// Mitsubishi GX Works2 project: AGV_IOCHECK   PLC: Q03UD

PROGRAM IOCHECK
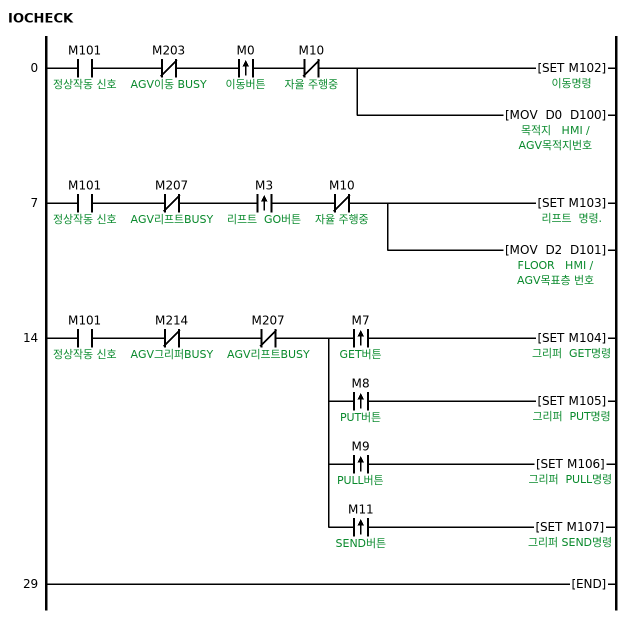
0     LD      M101  ; 정상작동 신호
      ANI     M203  ; AGV이동 BUSY
      ANDP    M0  ; 이동버튼
      ANI     M10  ; 자율 주행중
      SET     M102  ; 이동명령
      MOV     D0 D100  ; 목적지   HMI / AGV목적지번호
7     LD      M101  ; 정상작동 신호
      ANI     M207  ; AGV리프트BUSY
      ANDP    M3  ; 리프트  GO버튼
      ANI     M10  ; 자율 주행중
      SET     M103  ; 리프트  명령.
      MOV     D2 D101  ; FLOOR   HMI / AGV목표층 번호
14    LD      M101  ; 정상작동 신호
      ANI     M214  ; AGV그리퍼BUSY
      ANI     M207  ; AGV리프트BUSY
      MPS
      ANDP    M7  ; GET버튼
      SET     M104  ; 그리퍼  GET명령
      MRD
      ANDP    M8  ; PUT버튼
      SET     M105  ; 그리퍼  PUT명령
      MRD
      ANDP    M9  ; PULL버튼
      SET     M106  ; 그리퍼  PULL명령
      MPP
      ANDP    M11  ; SEND버튼
      SET     M107  ; 그리퍼 SEND명령
29    END
END_PROGRAM

PROGRAM MAIN
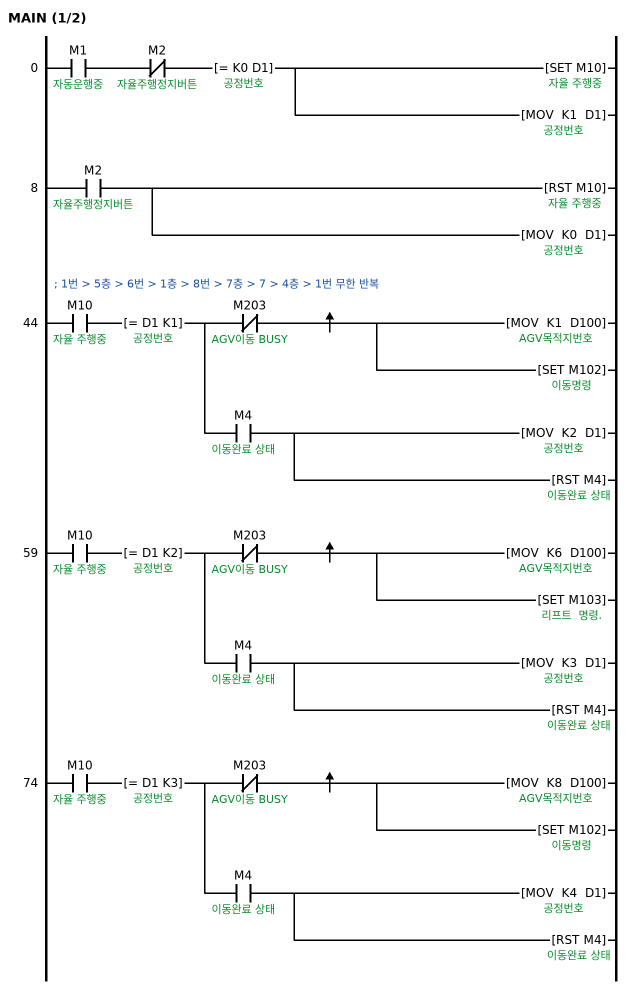
0     LD      M1  ; 자동운행중
      ANI     M2  ; 자율주행정지버튼
      AND=    K0 D1  ; 공정번호
      SET     M10  ; 자율 주행중
      MOV     K1 D1
8     LD      M2  ; 자율주행정지버튼
      RST     M10  ; 자율 주행중
      MOV     K0 D1
; 1번 > 5층 > 6번 > 1층 > 8번 > 7층 > 7 > 4층 > 1번 무한 반복
44    LD      M10  ; 자율 주행중
      AND=    D1 K1  ; 공정번호
      MPS
      ANI     M203  ; AGV이동 BUSY
      MEP
      MOV     K1 D100  ; AGV목적지번호
      SET     M102  ; 이동명령
      MPP
      AND     M4  ; 이동완료 상태
      MOV     K2 D1
      RST     M4  ; 이동완료 상태
59    LD      M10  ; 자율 주행중
      AND=    D1 K2  ; 공정번호
      MPS
      ANI     M203  ; AGV이동 BUSY
      MEP
      MOV     K6 D100
      SET     M103  ; 리프트  명령.
      MPP
      AND     M4  ; 이동완료 상태
      MOV     K3 D1
      RST     M4  ; 이동완료 상태
74    LD      M10  ; 자율 주행중
      AND=    D1 K3  ; 공정번호
      MPS
      ANI     M203  ; AGV이동 BUSY
      MEP
      MOV     K8 D100
      SET     M102  ; 이동명령
      MPP
      AND     M4  ; 이동완료 상태
      MOV     K4 D1
      RST     M4  ; 이동완료 상태
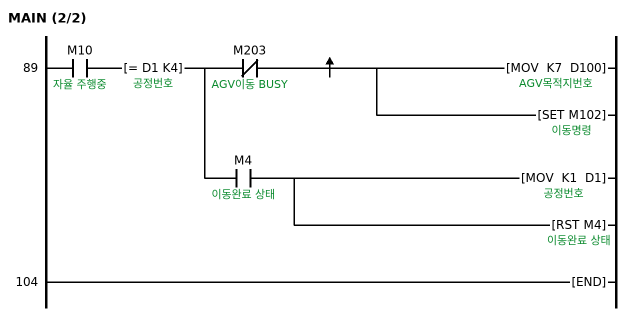
89    LD      M10  ; 자율 주행중
      AND=    D1 K4  ; 공정번호
      MPS
      ANI     M203  ; AGV이동 BUSY
      MEP
      MOV     K7 D100
      SET     M102  ; 이동명령
      MPP
      AND     M4  ; 이동완료 상태
      MOV     K1 D1
      RST     M4  ; 이동완료 상태
104   END
END_PROGRAM

PROGRAM MAIN2
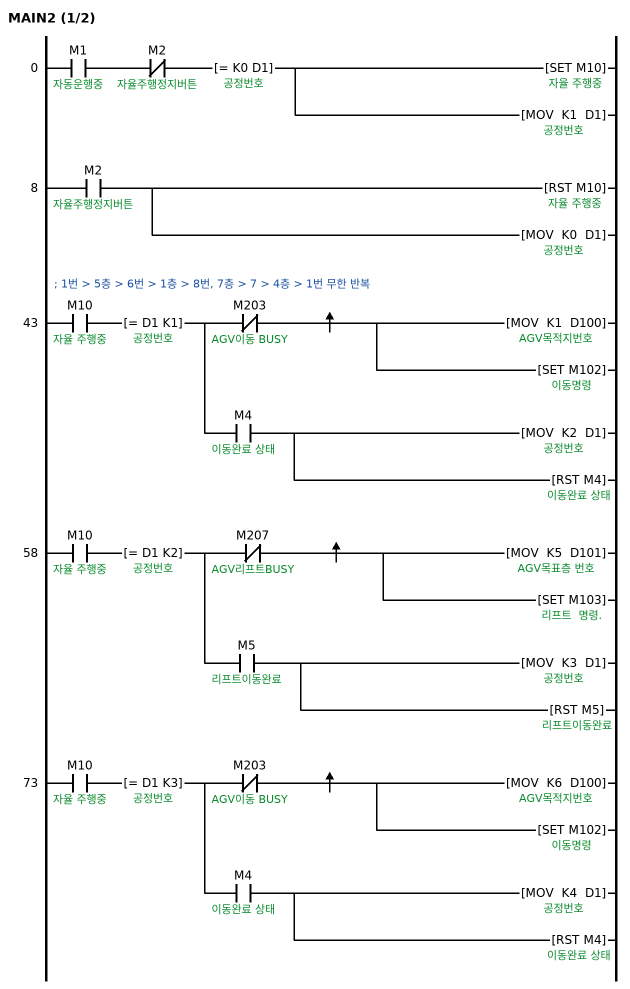
0     LD      M1  ; 자동운행중
      ANI     M2  ; 자율주행정지버튼
      AND=    K0 D1  ; 공정번호
      SET     M10  ; 자율 주행중
      MOV     K1 D1
8     LD      M2  ; 자율주행정지버튼
      RST     M10  ; 자율 주행중
      MOV     K0 D1
; 1번 > 5층 > 6번 > 1층 > 8번, 7층 > 7 > 4층 > 1번 무한 반복
43    LD      M10  ; 자율 주행중
      AND=    D1 K1  ; 공정번호
      MPS
      ANI     M203  ; AGV이동 BUSY
      MEP
      MOV     K1 D100  ; AGV목적지번호
      SET     M102  ; 이동명령
      MPP
      AND     M4  ; 이동완료 상태
      MOV     K2 D1
      RST     M4  ; 이동완료 상태
58    LD      M10  ; 자율 주행중
      AND=    D1 K2  ; 공정번호
      MPS
      ANI     M207  ; AGV리프트BUSY
      MEP
      MOV     K5 D101  ; AGV목표층 번호
      SET     M103  ; 리프트  명령.
      MPP
      AND     M5  ; 리프트이동완료
      MOV     K3 D1
      RST     M5  ; 리프트이동완료
73    LD      M10  ; 자율 주행중
      AND=    D1 K3  ; 공정번호
      MPS
      ANI     M203  ; AGV이동 BUSY
      MEP
      MOV     K6 D100
      SET     M102  ; 이동명령
      MPP
      AND     M4  ; 이동완료 상태
      MOV     K4 D1
      RST     M4  ; 이동완료 상태
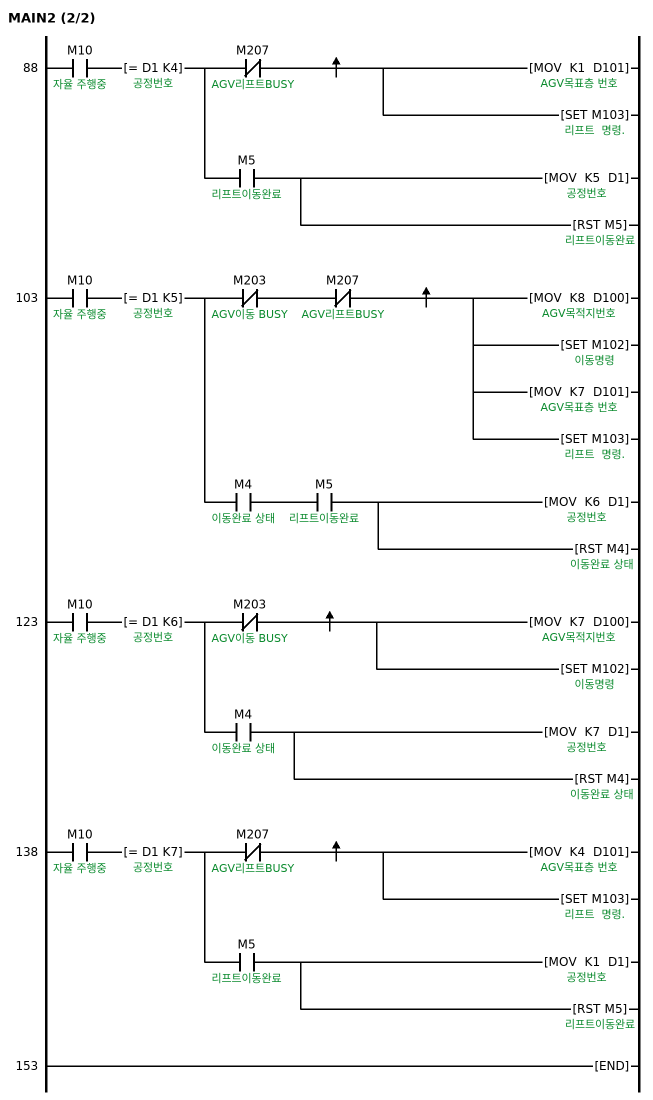
88    LD      M10  ; 자율 주행중
      AND=    D1 K4  ; 공정번호
      MPS
      ANI     M207  ; AGV리프트BUSY
      MEP
      MOV     K1 D101
      SET     M103  ; 리프트  명령.
      MPP
      AND     M5  ; 리프트이동완료
      MOV     K5 D1
      RST     M5  ; 리프트이동완료
103   LD      M10  ; 자율 주행중
      AND=    D1 K5  ; 공정번호
      MPS
      ANI     M203  ; AGV이동 BUSY
      ANI     M207  ; AGV리프트BUSY
      MEP
      MOV     K8 D100
      SET     M102  ; 이동명령
      MOV     K7 D101
      SET     M103  ; 리프트  명령.
      MPP
      AND     M4  ; 이동완료 상태
      AND     M5  ; 리프트이동완료
      MOV     K6 D1
      RST     M4  ; 이동완료 상태
123   LD      M10  ; 자율 주행중
      AND=    D1 K6  ; 공정번호
      MPS
      ANI     M203  ; AGV이동 BUSY
      MEP
      MOV     K7 D100
      SET     M102  ; 이동명령
      MPP
      AND     M4  ; 이동완료 상태
      MOV     K7 D1
      RST     M4  ; 이동완료 상태
138   LD      M10  ; 자율 주행중
      AND=    D1 K7  ; 공정번호
      MPS
      ANI     M207  ; AGV리프트BUSY
      MEP
      MOV     K4 D101
      SET     M103  ; 리프트  명령.
      MPP
      AND     M5  ; 리프트이동완료
      MOV     K1 D1
      RST     M5  ; 리프트이동완료
153   END
END_PROGRAM

PROGRAM INPUT
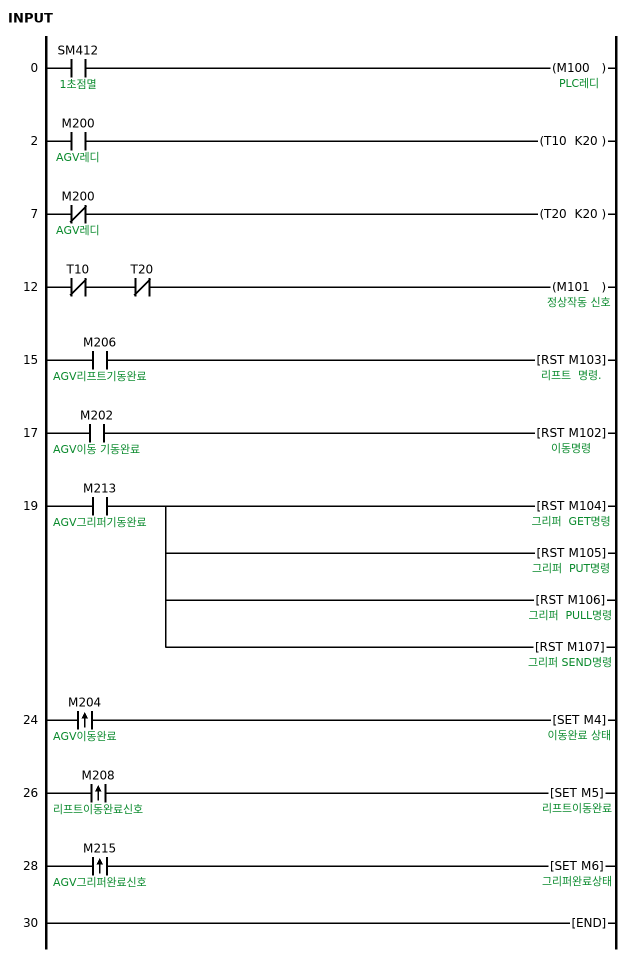
0     LD      SM412  ; 1초점멸
      OUT     M100  ; PLC레디
2     LD      M200  ; AGV레디
      OUT     T10 K20
7     LDI     M200  ; AGV레디
      OUT     T20 K20
12    LDI     T10
      ANI     T20
      OUT     M101  ; 정상작동 신호
15    LD      M206  ; AGV리프트기동완료
      RST     M103  ; 리프트  명령.
17    LD      M202  ; AGV이동 기동완료
      RST     M102  ; 이동명령
19    LD      M213  ; AGV그리퍼기동완료
      RST     M104  ; 그리퍼  GET명령
      RST     M105  ; 그리퍼  PUT명령
      RST     M106  ; 그리퍼  PULL명령
      RST     M107  ; 그리퍼 SEND명령
24    LDP     M204  ; AGV이동완료
      SET     M4  ; 이동완료 상태
26    LDP     M208  ; 리프트이동완료신호
      SET     M5  ; 리프트이동완료
28    LDP     M215  ; AGV그리퍼완료신호
      SET     M6  ; 그리퍼완료상태
30    END
END_PROGRAM

PROGRAM OUTPUT
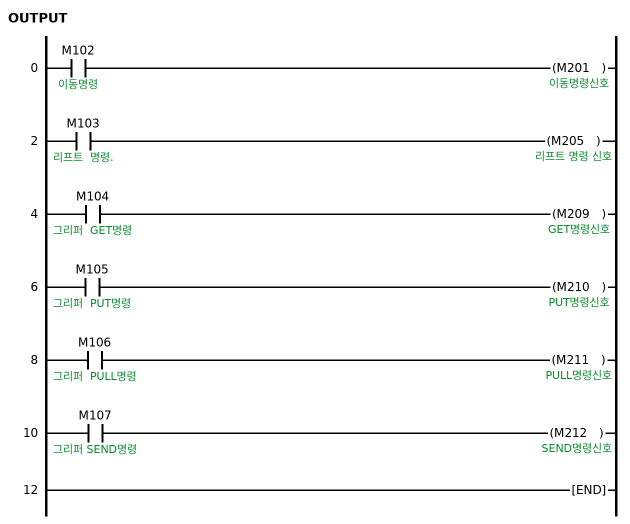
0     LD      M102  ; 이동명령
      OUT     M201  ; 이동명령신호
2     LD      M103  ; 리프트  명령.
      OUT     M205  ; 리프트 명령 신호
4     LD      M104  ; 그리퍼  GET명령
      OUT     M209  ; GET명령신호
6     LD      M105  ; 그리퍼  PUT명령
      OUT     M210  ; PUT명령신호
8     LD      M106  ; 그리퍼  PULL명령
      OUT     M211  ; PULL명령신호
10    LD      M107  ; 그리퍼 SEND명령
      OUT     M212  ; SEND명령신호
12    END
END_PROGRAM

PROGRAM MAIN3
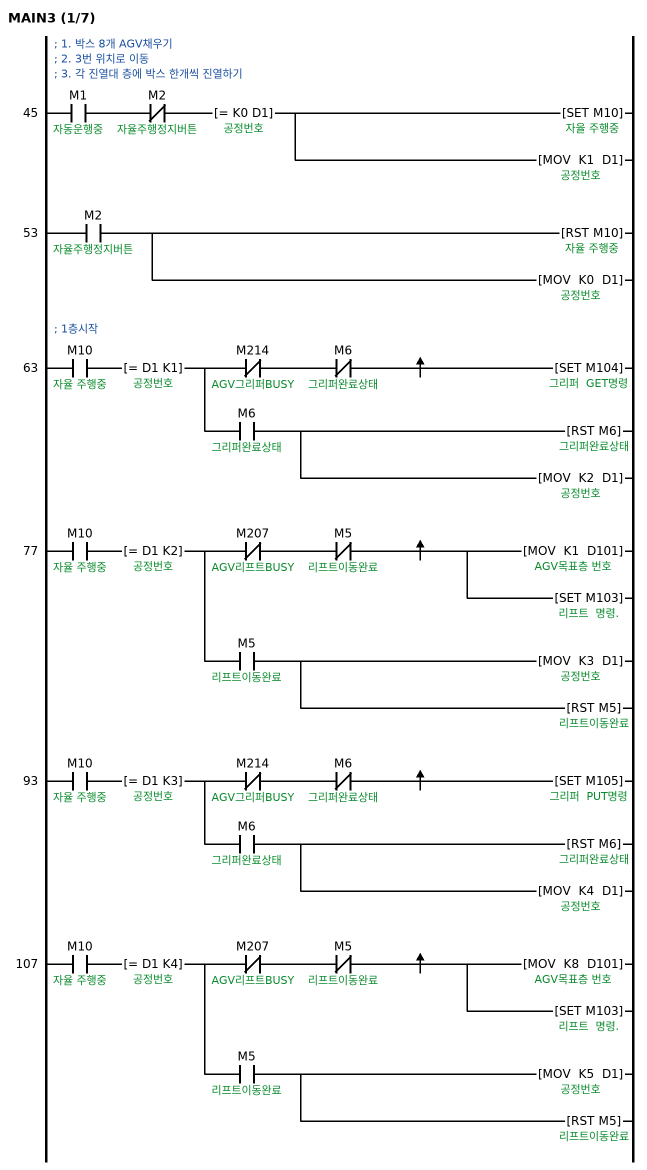
; 1. 박스 8개 AGV채우기
; 2. 3번 위치로 이동
; 3. 각 진열대 층에 박스 한개씩 진열하기
45    LD      M1  ; 자동운행중
      ANI     M2  ; 자율주행정지버튼
      AND=    K0 D1  ; 공정번호
      SET     M10  ; 자율 주행중
      MOV     K1 D1
53    LD      M2  ; 자율주행정지버튼
      RST     M10  ; 자율 주행중
      MOV     K0 D1
; 1층시작
63    LD      M10  ; 자율 주행중
      AND=    D1 K1  ; 공정번호
      MPS
      ANI     M214  ; AGV그리퍼BUSY
      ANI     M6  ; 그리퍼완료상태
      MEP
      SET     M104  ; 그리퍼  GET명령
      MPP
      AND     M6  ; 그리퍼완료상태
      RST     M6  ; 그리퍼완료상태
      MOV     K2 D1
77    LD      M10  ; 자율 주행중
      AND=    D1 K2  ; 공정번호
      MPS
      ANI     M207  ; AGV리프트BUSY
      ANI     M5  ; 리프트이동완료
      MEP
      MOV     K1 D101  ; AGV목표층 번호
      SET     M103  ; 리프트  명령.
      MPP
      AND     M5  ; 리프트이동완료
      MOV     K3 D1
      RST     M5  ; 리프트이동완료
93    LD      M10  ; 자율 주행중
      AND=    D1 K3  ; 공정번호
      MPS
      ANI     M214  ; AGV그리퍼BUSY
      ANI     M6  ; 그리퍼완료상태
      MEP
      SET     M105  ; 그리퍼  PUT명령
      MPP
      AND     M6  ; 그리퍼완료상태
      RST     M6  ; 그리퍼완료상태
      MOV     K4 D1
107   LD      M10  ; 자율 주행중
      AND=    D1 K4  ; 공정번호
      MPS
      ANI     M207  ; AGV리프트BUSY
      ANI     M5  ; 리프트이동완료
      MEP
      MOV     K8 D101
      SET     M103  ; 리프트  명령.
      MPP
      AND     M5  ; 리프트이동완료
      MOV     K5 D1
      RST     M5  ; 리프트이동완료
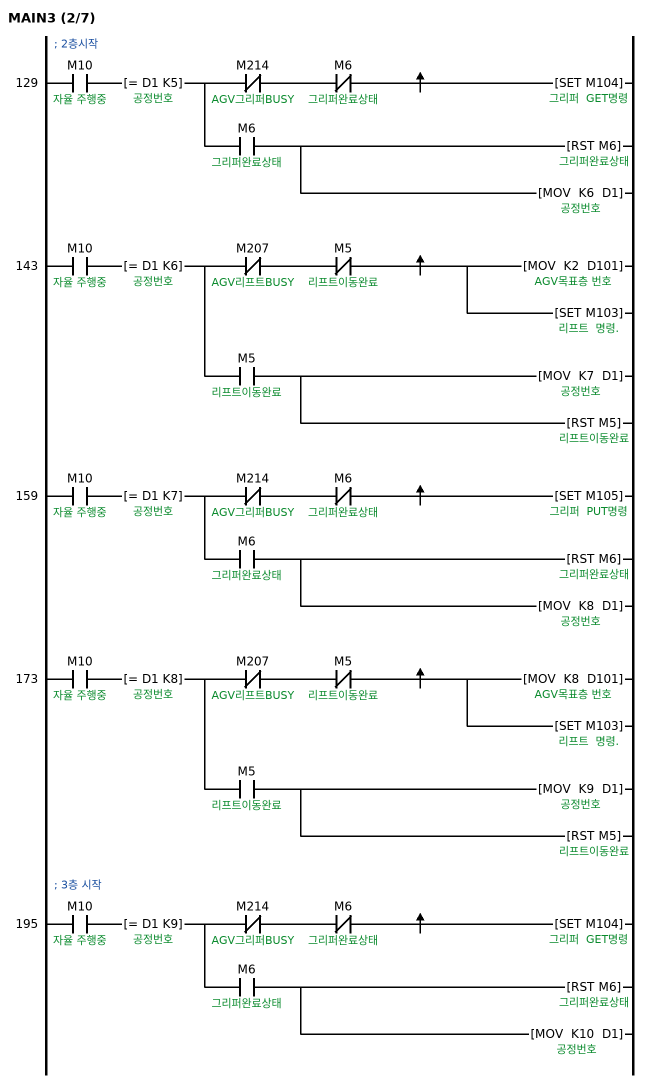
; 2층시작
129   LD      M10  ; 자율 주행중
      AND=    D1 K5  ; 공정번호
      MPS
      ANI     M214  ; AGV그리퍼BUSY
      ANI     M6  ; 그리퍼완료상태
      MEP
      SET     M104  ; 그리퍼  GET명령
      MPP
      AND     M6  ; 그리퍼완료상태
      RST     M6  ; 그리퍼완료상태
      MOV     K6 D1
143   LD      M10  ; 자율 주행중
      AND=    D1 K6  ; 공정번호
      MPS
      ANI     M207  ; AGV리프트BUSY
      ANI     M5  ; 리프트이동완료
      MEP
      MOV     K2 D101
      SET     M103  ; 리프트  명령.
      MPP
      AND     M5  ; 리프트이동완료
      MOV     K7 D1
      RST     M5  ; 리프트이동완료
159   LD      M10  ; 자율 주행중
      AND=    D1 K7  ; 공정번호
      MPS
      ANI     M214  ; AGV그리퍼BUSY
      ANI     M6  ; 그리퍼완료상태
      MEP
      SET     M105  ; 그리퍼  PUT명령
      MPP
      AND     M6  ; 그리퍼완료상태
      RST     M6  ; 그리퍼완료상태
      MOV     K8 D1
173   LD      M10  ; 자율 주행중
      AND=    D1 K8  ; 공정번호
      MPS
      ANI     M207  ; AGV리프트BUSY
      ANI     M5  ; 리프트이동완료
      MEP
      MOV     K8 D101
      SET     M103  ; 리프트  명령.
      MPP
      AND     M5  ; 리프트이동완료
      MOV     K9 D1
      RST     M5  ; 리프트이동완료
; 3층 시작
195   LD      M10  ; 자율 주행중
      AND=    D1 K9  ; 공정번호
      MPS
      ANI     M214  ; AGV그리퍼BUSY
      ANI     M6  ; 그리퍼완료상태
      MEP
      SET     M104  ; 그리퍼  GET명령
      MPP
      AND     M6  ; 그리퍼완료상태
      RST     M6  ; 그리퍼완료상태
      MOV     K10 D1
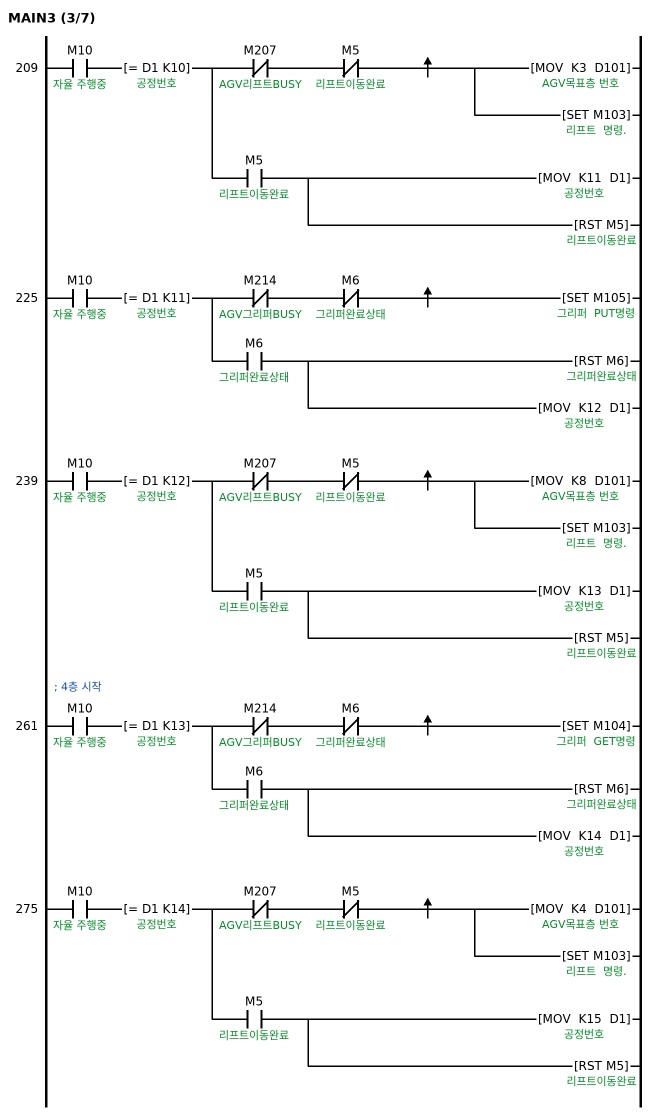
209   LD      M10  ; 자율 주행중
      AND=    D1 K10  ; 공정번호
      MPS
      ANI     M207  ; AGV리프트BUSY
      ANI     M5  ; 리프트이동완료
      MEP
      MOV     K3 D101
      SET     M103  ; 리프트  명령.
      MPP
      AND     M5  ; 리프트이동완료
      MOV     K11 D1
      RST     M5  ; 리프트이동완료
225   LD      M10  ; 자율 주행중
      AND=    D1 K11  ; 공정번호
      MPS
      ANI     M214  ; AGV그리퍼BUSY
      ANI     M6  ; 그리퍼완료상태
      MEP
      SET     M105  ; 그리퍼  PUT명령
      MPP
      AND     M6  ; 그리퍼완료상태
      RST     M6  ; 그리퍼완료상태
      MOV     K12 D1
239   LD      M10  ; 자율 주행중
      AND=    D1 K12  ; 공정번호
      MPS
      ANI     M207  ; AGV리프트BUSY
      ANI     M5  ; 리프트이동완료
      MEP
      MOV     K8 D101
      SET     M103  ; 리프트  명령.
      MPP
      AND     M5  ; 리프트이동완료
      MOV     K13 D1
      RST     M5  ; 리프트이동완료
; 4층 시작
261   LD      M10  ; 자율 주행중
      AND=    D1 K13  ; 공정번호
      MPS
      ANI     M214  ; AGV그리퍼BUSY
      ANI     M6  ; 그리퍼완료상태
      MEP
      SET     M104  ; 그리퍼  GET명령
      MPP
      AND     M6  ; 그리퍼완료상태
      RST     M6  ; 그리퍼완료상태
      MOV     K14 D1
275   LD      M10  ; 자율 주행중
      AND=    D1 K14  ; 공정번호
      MPS
      ANI     M207  ; AGV리프트BUSY
      ANI     M5  ; 리프트이동완료
      MEP
      MOV     K4 D101
      SET     M103  ; 리프트  명령.
      MPP
      AND     M5  ; 리프트이동완료
      MOV     K15 D1
      RST     M5  ; 리프트이동완료
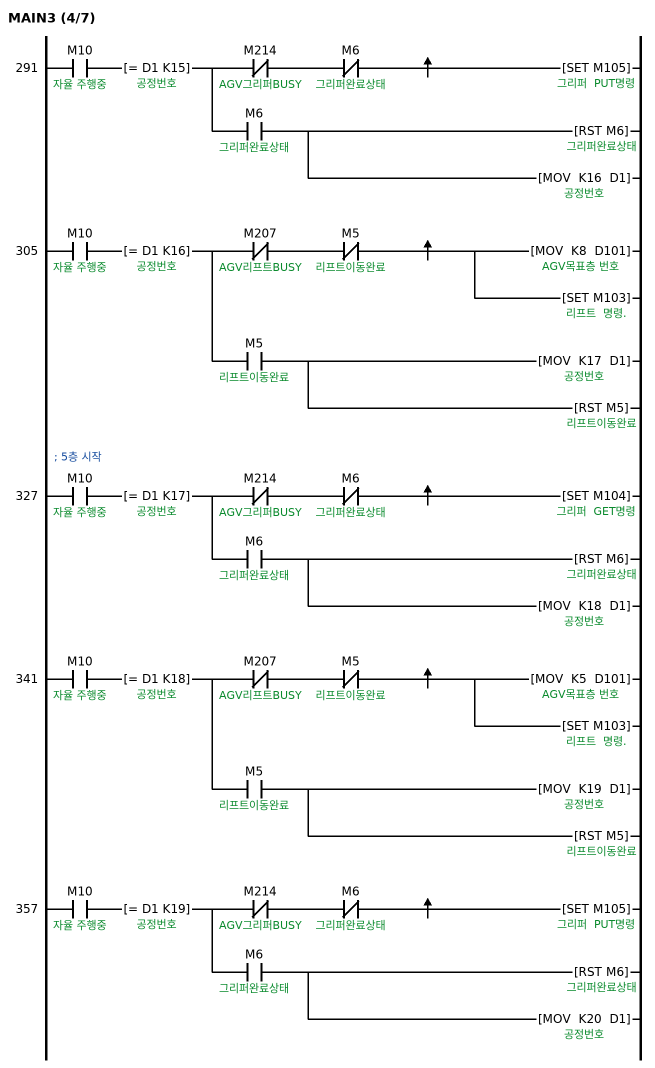
291   LD      M10  ; 자율 주행중
      AND=    D1 K15  ; 공정번호
      MPS
      ANI     M214  ; AGV그리퍼BUSY
      ANI     M6  ; 그리퍼완료상태
      MEP
      SET     M105  ; 그리퍼  PUT명령
      MPP
      AND     M6  ; 그리퍼완료상태
      RST     M6  ; 그리퍼완료상태
      MOV     K16 D1
305   LD      M10  ; 자율 주행중
      AND=    D1 K16  ; 공정번호
      MPS
      ANI     M207  ; AGV리프트BUSY
      ANI     M5  ; 리프트이동완료
      MEP
      MOV     K8 D101
      SET     M103  ; 리프트  명령.
      MPP
      AND     M5  ; 리프트이동완료
      MOV     K17 D1
      RST     M5  ; 리프트이동완료
; 5층 시작
327   LD      M10  ; 자율 주행중
      AND=    D1 K17  ; 공정번호
      MPS
      ANI     M214  ; AGV그리퍼BUSY
      ANI     M6  ; 그리퍼완료상태
      MEP
      SET     M104  ; 그리퍼  GET명령
      MPP
      AND     M6  ; 그리퍼완료상태
      RST     M6  ; 그리퍼완료상태
      MOV     K18 D1
341   LD      M10  ; 자율 주행중
      AND=    D1 K18  ; 공정번호
      MPS
      ANI     M207  ; AGV리프트BUSY
      ANI     M5  ; 리프트이동완료
      MEP
      MOV     K5 D101
      SET     M103  ; 리프트  명령.
      MPP
      AND     M5  ; 리프트이동완료
      MOV     K19 D1
      RST     M5  ; 리프트이동완료
357   LD      M10  ; 자율 주행중
      AND=    D1 K19  ; 공정번호
      MPS
      ANI     M214  ; AGV그리퍼BUSY
      ANI     M6  ; 그리퍼완료상태
      MEP
      SET     M105  ; 그리퍼  PUT명령
      MPP
      AND     M6  ; 그리퍼완료상태
      RST     M6  ; 그리퍼완료상태
      MOV     K20 D1
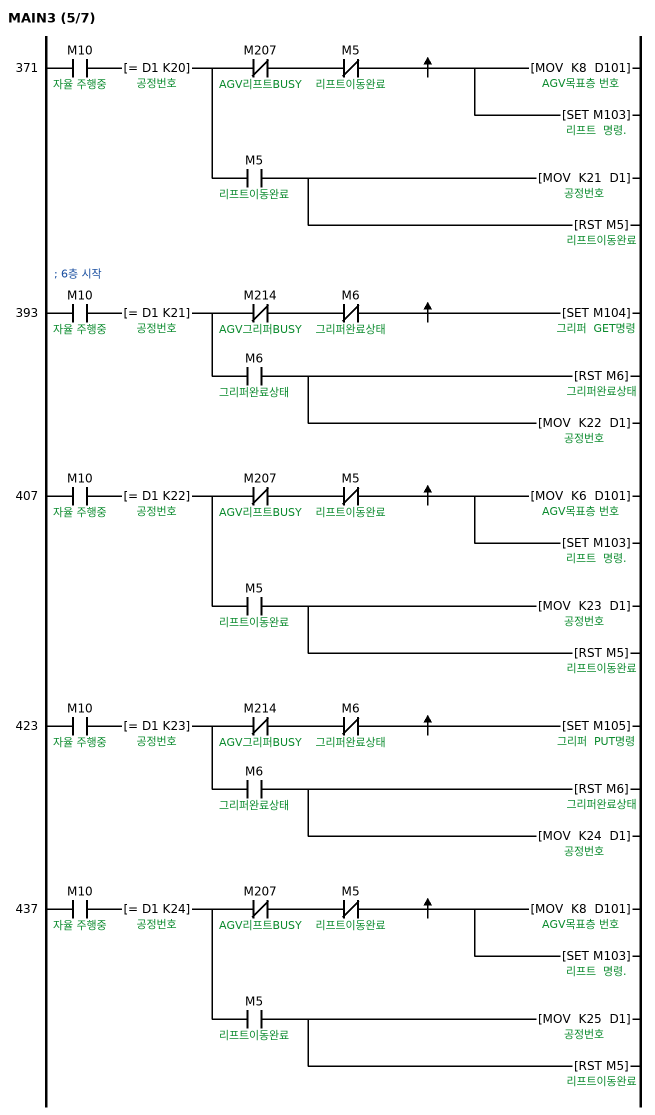
371   LD      M10  ; 자율 주행중
      AND=    D1 K20  ; 공정번호
      MPS
      ANI     M207  ; AGV리프트BUSY
      ANI     M5  ; 리프트이동완료
      MEP
      MOV     K8 D101
      SET     M103  ; 리프트  명령.
      MPP
      AND     M5  ; 리프트이동완료
      MOV     K21 D1
      RST     M5  ; 리프트이동완료
; 6층 시작
393   LD      M10  ; 자율 주행중
      AND=    D1 K21  ; 공정번호
      MPS
      ANI     M214  ; AGV그리퍼BUSY
      ANI     M6  ; 그리퍼완료상태
      MEP
      SET     M104  ; 그리퍼  GET명령
      MPP
      AND     M6  ; 그리퍼완료상태
      RST     M6  ; 그리퍼완료상태
      MOV     K22 D1
407   LD      M10  ; 자율 주행중
      AND=    D1 K22  ; 공정번호
      MPS
      ANI     M207  ; AGV리프트BUSY
      ANI     M5  ; 리프트이동완료
      MEP
      MOV     K6 D101
      SET     M103  ; 리프트  명령.
      MPP
      AND     M5  ; 리프트이동완료
      MOV     K23 D1
      RST     M5  ; 리프트이동완료
423   LD      M10  ; 자율 주행중
      AND=    D1 K23  ; 공정번호
      MPS
      ANI     M214  ; AGV그리퍼BUSY
      ANI     M6  ; 그리퍼완료상태
      MEP
      SET     M105  ; 그리퍼  PUT명령
      MPP
      AND     M6  ; 그리퍼완료상태
      RST     M6  ; 그리퍼완료상태
      MOV     K24 D1
437   LD      M10  ; 자율 주행중
      AND=    D1 K24  ; 공정번호
      MPS
      ANI     M207  ; AGV리프트BUSY
      ANI     M5  ; 리프트이동완료
      MEP
      MOV     K8 D101
      SET     M103  ; 리프트  명령.
      MPP
      AND     M5  ; 리프트이동완료
      MOV     K25 D1
      RST     M5  ; 리프트이동완료
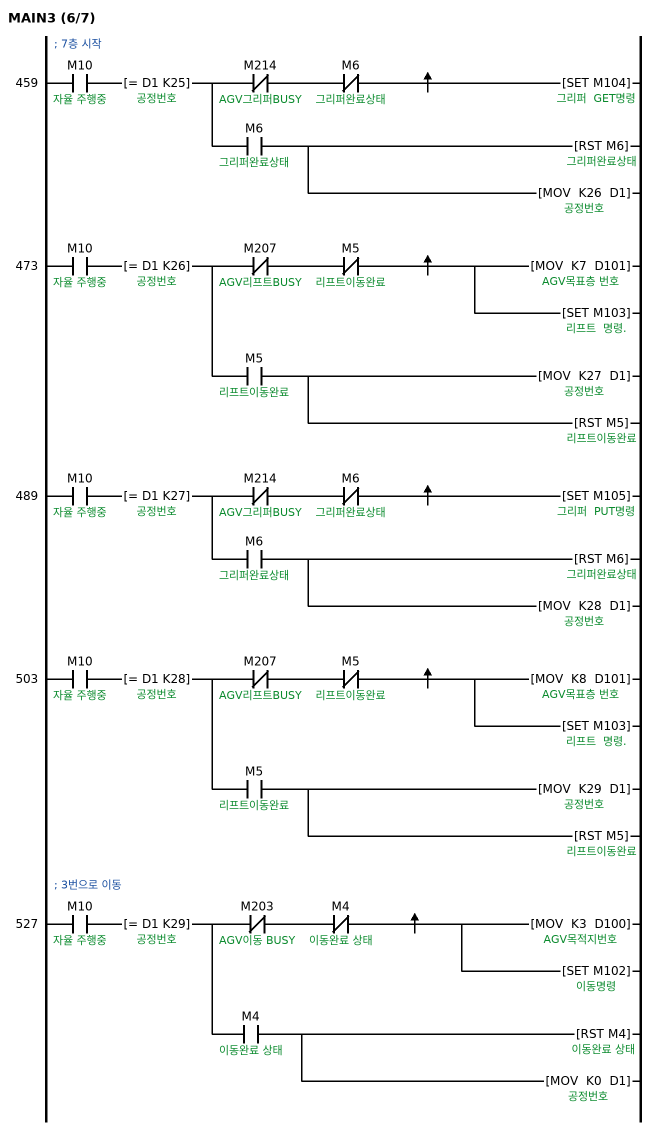
; 7층 시작
459   LD      M10  ; 자율 주행중
      AND=    D1 K25  ; 공정번호
      MPS
      ANI     M214  ; AGV그리퍼BUSY
      ANI     M6  ; 그리퍼완료상태
      MEP
      SET     M104  ; 그리퍼  GET명령
      MPP
      AND     M6  ; 그리퍼완료상태
      RST     M6  ; 그리퍼완료상태
      MOV     K26 D1
473   LD      M10  ; 자율 주행중
      AND=    D1 K26  ; 공정번호
      MPS
      ANI     M207  ; AGV리프트BUSY
      ANI     M5  ; 리프트이동완료
      MEP
      MOV     K7 D101
      SET     M103  ; 리프트  명령.
      MPP
      AND     M5  ; 리프트이동완료
      MOV     K27 D1
      RST     M5  ; 리프트이동완료
489   LD      M10  ; 자율 주행중
      AND=    D1 K27  ; 공정번호
      MPS
      ANI     M214  ; AGV그리퍼BUSY
      ANI     M6  ; 그리퍼완료상태
      MEP
      SET     M105  ; 그리퍼  PUT명령
      MPP
      AND     M6  ; 그리퍼완료상태
      RST     M6  ; 그리퍼완료상태
      MOV     K28 D1
503   LD      M10  ; 자율 주행중
      AND=    D1 K28  ; 공정번호
      MPS
      ANI     M207  ; AGV리프트BUSY
      ANI     M5  ; 리프트이동완료
      MEP
      MOV     K8 D101
      SET     M103  ; 리프트  명령.
      MPP
      AND     M5  ; 리프트이동완료
      MOV     K29 D1
      RST     M5  ; 리프트이동완료
; 3번으로 이동
527   LD      M10  ; 자율 주행중
      AND=    D1 K29  ; 공정번호
      MPS
      ANI     M203  ; AGV이동 BUSY
      ANI     M4  ; 이동완료 상태
      MEP
      MOV     K3 D100  ; AGV목적지번호
      SET     M102  ; 이동명령
      MPP
      AND     M4  ; 이동완료 상태
      RST     M4  ; 이동완료 상태
      MOV     K0 D1
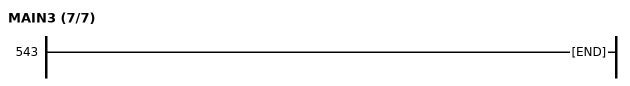
543   END
END_PROGRAM

PROGRAM TEST
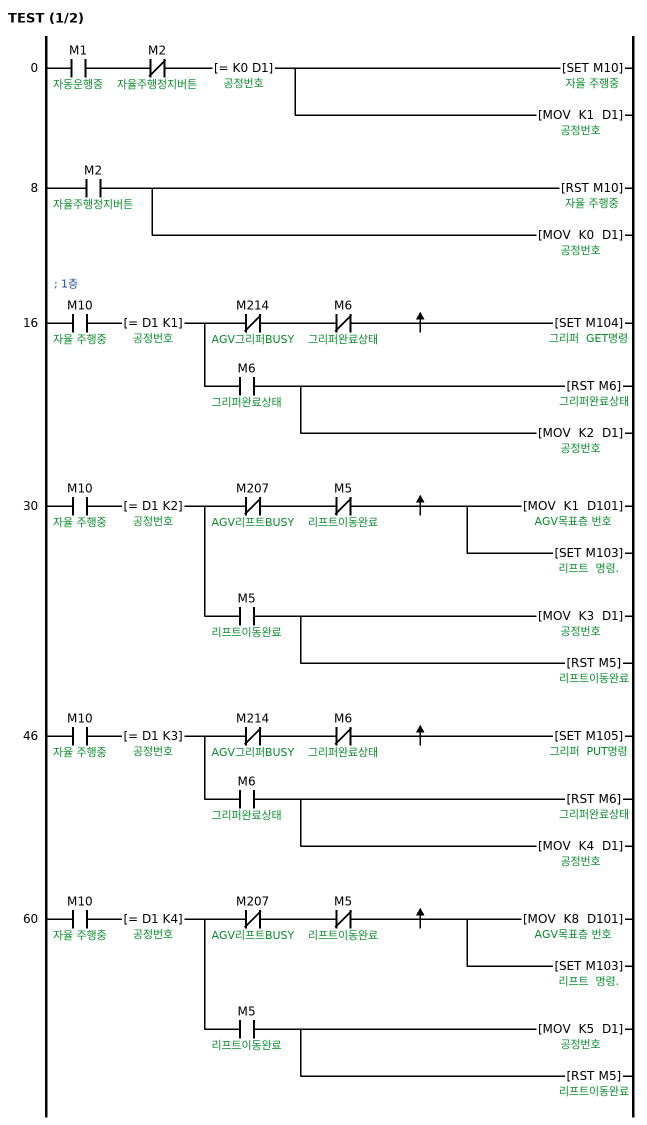
0     LD      M1  ; 자동운행중
      ANI     M2  ; 자율주행정지버튼
      AND=    K0 D1  ; 공정번호
      SET     M10  ; 자율 주행중
      MOV     K1 D1
8     LD      M2  ; 자율주행정지버튼
      RST     M10  ; 자율 주행중
      MOV     K0 D1
; 1층
16    LD      M10  ; 자율 주행중
      AND=    D1 K1  ; 공정번호
      MPS
      ANI     M214  ; AGV그리퍼BUSY
      ANI     M6  ; 그리퍼완료상태
      MEP
      SET     M104  ; 그리퍼  GET명령
      MPP
      AND     M6  ; 그리퍼완료상태
      RST     M6  ; 그리퍼완료상태
      MOV     K2 D1
30    LD      M10  ; 자율 주행중
      AND=    D1 K2  ; 공정번호
      MPS
      ANI     M207  ; AGV리프트BUSY
      ANI     M5  ; 리프트이동완료
      MEP
      MOV     K1 D101  ; AGV목표층 번호
      SET     M103  ; 리프트  명령.
      MPP
      AND     M5  ; 리프트이동완료
      MOV     K3 D1
      RST     M5  ; 리프트이동완료
46    LD      M10  ; 자율 주행중
      AND=    D1 K3  ; 공정번호
      MPS
      ANI     M214  ; AGV그리퍼BUSY
      ANI     M6  ; 그리퍼완료상태
      MEP
      SET     M105  ; 그리퍼  PUT명령
      MPP
      AND     M6  ; 그리퍼완료상태
      RST     M6  ; 그리퍼완료상태
      MOV     K4 D1
60    LD      M10  ; 자율 주행중
      AND=    D1 K4  ; 공정번호
      MPS
      ANI     M207  ; AGV리프트BUSY
      ANI     M5  ; 리프트이동완료
      MEP
      MOV     K8 D101
      SET     M103  ; 리프트  명령.
      MPP
      AND     M5  ; 리프트이동완료
      MOV     K5 D1
      RST     M5  ; 리프트이동완료
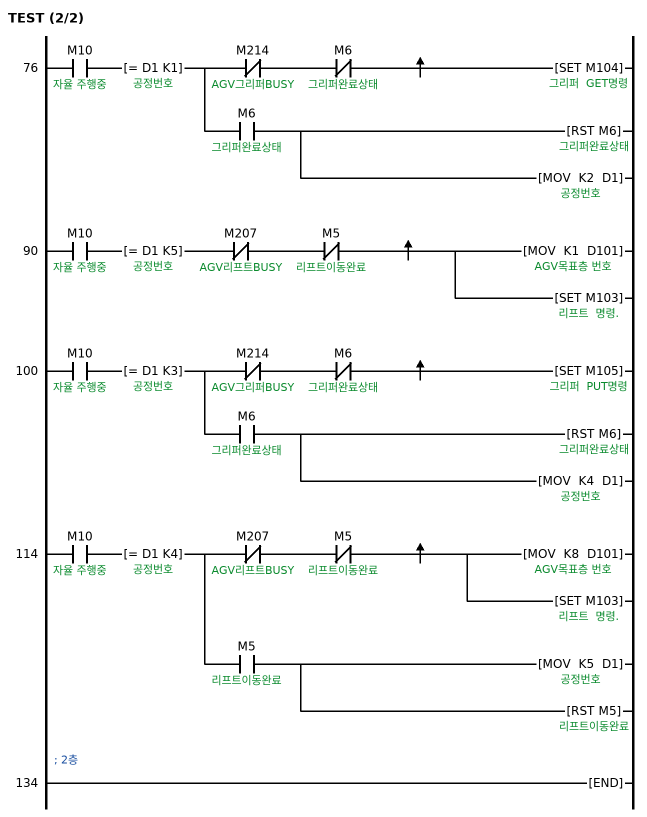
76    LD      M10  ; 자율 주행중
      AND=    D1 K1  ; 공정번호
      MPS
      ANI     M214  ; AGV그리퍼BUSY
      ANI     M6  ; 그리퍼완료상태
      MEP
      SET     M104  ; 그리퍼  GET명령
      MPP
      AND     M6  ; 그리퍼완료상태
      RST     M6  ; 그리퍼완료상태
      MOV     K2 D1
90    LD      M10  ; 자율 주행중
      AND=    D1 K5  ; 공정번호
      ANI     M207  ; AGV리프트BUSY
      ANI     M5  ; 리프트이동완료
      MEP
      MOV     K1 D101
      SET     M103  ; 리프트  명령.
100   LD      M10  ; 자율 주행중
      AND=    D1 K3  ; 공정번호
      MPS
      ANI     M214  ; AGV그리퍼BUSY
      ANI     M6  ; 그리퍼완료상태
      MEP
      SET     M105  ; 그리퍼  PUT명령
      MPP
      AND     M6  ; 그리퍼완료상태
      RST     M6  ; 그리퍼완료상태
      MOV     K4 D1
114   LD      M10  ; 자율 주행중
      AND=    D1 K4  ; 공정번호
      MPS
      ANI     M207  ; AGV리프트BUSY
      ANI     M5  ; 리프트이동완료
      MEP
      MOV     K8 D101
      SET     M103  ; 리프트  명령.
      MPP
      AND     M5  ; 리프트이동완료
      MOV     K5 D1
      RST     M5  ; 리프트이동완료
; 2층
134   END
END_PROGRAM

PROGRAM FINAL
0     END
END_PROGRAM

// device comments not shown above
Y20  ; 반복
Y40  ; GET
Y41  ; GET
Y42  ; RESET
Y43  ; PUT
